// TIA Portal V19 export
// export: Created 2026-11-02T08:00:00.000Z, ExportSetting WithDefaults
FUNCTION_BLOCK "FB_Conveyor"   // FB10, LAD
TITLE = Belt conveyor
{ S7_Optimized_Access := 'TRUE' }
AUTHOR : controls
VERSION : 0.1
// stored: AutoNumber true, SetENOAutomatically false
   VAR_INPUT
      Start : Bool;   // Start push button
      Stop : Bool;   // Stop push button
   END_VAR
   VAR_OUTPUT
      Run : Bool;
      JamAlarm : Bool;
   END_VAR
   VAR
      JamTimer : IEC_TIMER;
      Speed : Real := 1.2;
   END_VAR
BEGIN

REGION Network 1: Run latch
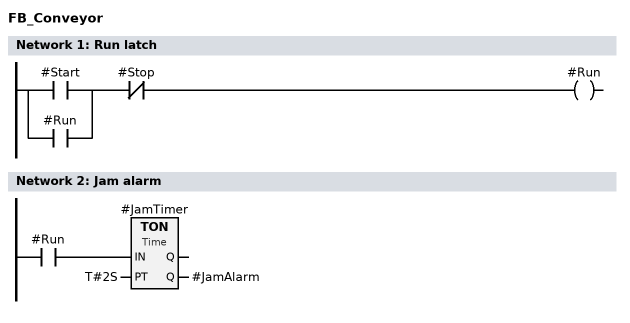
   RUNG wire#powerrail
      Contact( #Start )
      wire#w1
      I_Contact( #Stop )
      Coil( #Run )
   END_RUNG
   RUNG wire#powerrail
      Contact( #Run )
   END_RUNG wire#w1
   // the same network as SCL:
   #Run := (#Start OR #Run) AND NOT #Stop;
END_REGION

REGION Network 2: Jam alarm
   RUNG wire#powerrail
      Contact( #Run )
      { S7_Templates := "time_type := Time" } #JamTimer.TON(pt := T#2S, q => #JamAlarm)
   END_RUNG
   // the same network as SCL:
   #JamTimer.TON(IN := #Run, PT := T#2S, Q => #JamAlarm);
END_REGION
END_FUNCTION_BLOCK
